Fanuc KAREL source: kt00373.KL

-- PROVISIONAL review KL for V770-1; original PC SHA256 2e54453345df820f799d1481306cd7edc94904fc5b24947b02e420b27f0f7298
-- Incomplete behavior may be omitted. Consult companion uncertainty JSON. Do not deploy.
PROGRAM KT00373
%NOLOCKGROUP
VAR
  B1 : BOOLEAN
  B2 : BOOLEAN
  OUT : BOOLEAN
BEGIN
  -- UNRESOLVED_PC offsets 5-12; opcodes 9D,23
  -- UNRESOLVED_PC offsets 17-24; opcodes 9C,23
  -- UNRESOLVED_PC offsets 29-36; opcodes 9D,23
  -- UNRESOLVED_PC offsets 41-48; opcodes 9C,23
  -- UNRESOLVED_PC offsets 53-72; opcodes 21,21,5A,23
  -- UNRESOLVED_PC offsets 77-81; opcodes 7F
END KT00373
